(* IEC 61131-3 sources: volt/packages/volt-lsp-iec/test-corpus/awa-palletizer/Device/Plc Logic/Application/Library Manager/L_IPAP_ParameterManagerAccess, 29 files *)

(* ---- L_IPAP_DATATYPE.dut ---- *)
TYPE L_IPAP_DATATYPE :
(
	DT_EMPTY := 0,
	DT_STRING := 1,
	DT_WSTRING := 2,
	DT_BOOLEAN := 3,
	DT_INTEGER_8 := 4,
	DT_INTEGER_16 := 5,
	DT_INTEGER_32 := 6,
	DT_INTEGER_64 := 7,
	DT_UNSIGNED_8 := 8,
	DT_UNSIGNED_16 := 9,
	DT_UNSIGNED_32 := 10,
	DT_UNSIGNED_64 := 11,
	DT_FLOAT_32 := 12,
	DT_FLOAT_64 := 13,
	DT_OCTETSTRING := 14
);
END_TYPE

(* ---- L_IPAP_ERRORID.dut ---- *)
TYPE L_IPAP_ERRORID :
(
	ERR_NOERROR := 0,
	ERR_PARAMETERERROR,
	ERR_INTERNALERROR,
	ERR_TIMEOUT,
	ERR_PARAMETERNOTEXISTING,
	ERR_READACCESSDENIED,
	ERR_WRITEACCESSDENIED,
	ERR_VALUESIZEEXCEEDED,
	ERR_LOWLIMITVIOLATION,
	ERR_HIGHLIMITVIOLATION,
	ERR_NOSELECTLISTVALUE,
	ERR_CONTROLLERINHIBIT,
	ERR_BUFFERSIZE,
	ERR_HAPROXYNOTACTIVE,
	ERR_CHANGEHTTPSREDIRECTFAILED
);
END_TYPE

(* ---- L_IPAP_FBSTATE.dut ---- *)
TYPE L_IPAP_FBSTATE :
(
	INIT := 0,
	WAIT,
	START,
	CHECK,
	DONE,
	ERROR,
	ABORT,
	RESET,
	READ,
	WRITE,
	VERIFY
);
END_TYPE

(* ---- L_IPAP_HTTPSREDIRECT.dut ---- *)
TYPE L_IPAP_HTTPSREDIRECT :
(
	DISABLE_HTTPSREDIRECT := 0,
	ENABLE_HTTPSREDIRECT := 1
);
END_TYPE

(* ---- L_IPAP_INTERNALERROR.dut ---- *)
TYPE L_IPAP_INTERNALERROR :
(
	ERR_OK := 16#0,
	ERR_PROTOCOL_TIMEOUT := 16#2,
	ERR_OUT_OF_MEMORY := 16#4,
	ERR_UNSUPPORTED_ACCESS := 16#5,
	ERR_WRITE_ONLY_ENTRY := 16#6,
	ERR_READ_ONLY_ENTRY := 16#7,
	ERR_OBJECT_NOT_EXISTING := 16#8,
	ERR_PARAM_IS_INCOMPATIBLE := 16#B,
	ERR_INTERNAL_DEVICE_INCOMPATIBILITY := 16#C,
	ERR_PARAM_LENGTH_ERROR := 16#E,
	ERR_PARAM_LENGTH_TOO_LONG := 16#F,
	ERR_PARAM_LENGTH_TOO_SHORT := 16#10,
	ERR_SUBINDEX_NOT_EXISTING := 16#11,
	ERR_VALUE_EXCEEDED := 16#12,
	ERR_VALUE_TOO_GREAT := 16#13,
	ERR_VALUE_TOO_SMALL := 16#14,
	ERR_MAX_VALUE_IS_LESS_THAN_MIN_VALUE := 16#15,
	ERR_GENERAL_ERROR := 16#16,
	ERR_DATA_CANNOT_BE_READ_OR_STORED := 16#17,
	ERR_DATA_CANNOT_BE_READ_OR_STORED_BECAUSE_OF_LOCAL_CONTROL := 16#18,
	ERR_DATA_CANNOT_BE_READ_OR_STORED_IN_THIS_STATE := 16#19,
	ERR_SEND_REQUEST_FAILED := 16#50,
	ERR_UNKNOWN_DATATYPE := 16#51,
	ERR_BUFFER_SIZE := 16#52
);
END_TYPE

(* ---- L_IPAP_INTERNALERROR_ABORTCODE.dut ---- *)
TYPE L_IPAP_INTERNALERROR_ABORTCODE :
(
	ABORT_NOERROR := 16#0,
	ABORT_TIMEOUT := 16#5040000,
	ABORT_OUT_OF_MEMORY := 16#5040005,
	ABORT_UNSUPPORTED_ACCESS := 16#6010000,
	ABORT_WRITE_ONLY_ENTRY := 16#6010001,
	ABORT_READ_ONLY_ENTRY := 16#6010002,
	ABORT_OBJECT_NOT_EXISTING := 16#6020000,
	ABORT_PARAM_IS_INCOMPATIBLE := 16#6040043,
	ABORT_INTERNAL_DEVICE_INCOMPATIBILITY := 16#6040047,
	ABORT_PARAM_LENGTH_ERROR := 16#6070010,
	ABORT_PARAM_LENGTH_TOO_LONG := 16#6070012,
	ABORT_PARAM_LENGTH_TOO_SHORT := 16#6070013,
	ABORT_SUBINDEX_NOT_EXISTING := 16#6090011,
	ABORT_VALUE_EXCEEDED := 16#6090030,
	ABORT_VALUE_TOO_GREAT := 16#6090031,
	ABORT_VALUE_TOO_SMALL := 16#6090032,
	ABORT_MAX_VALUE_IS_LESS_THAN_MIN_VALUE := 16#6090036,
	ABORT_GENERAL_ERROR := 16#8000000,
	ABORT_DATA_CANNOT_BE_READ_OR_STORED := 16#8000020,
	ABORT_DATA_CANNOT_BE_READ_OR_STORED_BECAUSE_OF_LOCAL_CONTROL := 16#8000021,
	ABORT_DATA_CANNOT_BE_READ_OR_STORED_IN_THIS_STATE := 16#8000022
);
END_TYPE

(* ---- L_IPAP_INTERNALERROR_OLD.dut ---- *)
TYPE L_IPAP_INTERNALERROR_OLD :
(
	PMA_OK := 0,
	PMA_TOGGLEBITNOTCHANGED := 1,
	PMA_SDOPROTOCOLTIMEOUT := 2,
	PMA_COMMANDSPECIFIERUNKNOWN := 3,
	PMA_OUTOFMEMORY := 4,
	PMA_UNSUPPORTEDACCESS := 5,
	PMA_WRITEONLYENTRY := 6,
	PMA_READONLYENTRY := 7,
	PMA_OBJECTNOTEXISTING := 8,
	PMA_OBJECTCANTBEPDOMAPPED := 9,
	PMA_MAPPEDOBJECTSEXCEEDPDO := 10,
	PMA_PARAMISINCOMPATIBLE := 11,
	PMA_INTERNALDEVICEINCOMPATIBILITY := 12,
	PMA_HARDWAREERROR := 13,
	PMA_PARAMLENGTHERROR := 14,
	PMA_PARAMLENGTHTOOLONG := 15,
	PMA_PARAMLENGTHTOOSHORT := 16,
	PMA_SUBINDEXNOTEXISTING := 17,
	PMA_VALUEEXCEEDED := 18,
	PMA_VALUETOOGREAT := 19,
	PMA_VALUETOOSMALL := 20,
	PMA_MAXVALUEISLESSTHANMINVALUE := 21,
	PMA_GENERALERROR := 22,
	PMA_DATACANNOTBEREADORSTORED := 23,
	PMA_DATACANNOTBEACCESSEDBECAUSEOFLOCALCONTROL := 24,
	PMA_INTHISSTATEDATACANNOTBEREADORSTORED := 25,
	PMA_NOOBJECTDICTIONARYISPRESENT := 26,
	PMA_ENTRYCANTBEWRITTENSI0NOT0 := 27,
	PMA_COMPLETEACCESSNOTSUPPORTEDFFORTHISOBJ := 28,
	PMA_OBJLENGTHEXCEEDSMBXSIZE := 29,
	PMA_OBJMAPPEDTOPDOSDOACCESSBLOCKED := 30,
	PMA_BUFFEROVERFLOW := 33,
	PMA_INVALIDREPLY := 34,
	PMA_UNKNOWNCOMMAND := 35,
	PMA_PARAMETERERROR := 37,
	PMA_REPLYERROR := 38,
	PMA_REPLYTIMEOUT := 39,
	PMA_SERVERQUEUEERROR := 40,
	PMA_PROTOCOLMISMATCH := 41,
	PMA_SENDREQUESTFAILED := 70,
	PMA_UNKNOWNDATATYPE := 71,
	PMA_OTHERERROR := 99
);
END_TYPE

(* ---- L_IPAP_REQUEST_STATE.dut ---- *)
TYPE L_IPAP_REQUEST_STATE :
(
	UNKNOWN := 0,
	ERROR := 1,
	WAIT := 2,
	BUSY := 3,
	DONE := 4
);
END_TYPE

(* ---- GETBOOLEANPROPERTY.pou ---- *)
FUNCTION GETBOOLEANPROPERTY : BOOL
VAR_INPUT
	STKEY : WSTRING;
END_VAR
END_FUNCTION

(* ---- GETCOMPANY.pou ---- *)
FUNCTION GETCOMPANY : WSTRING
END_FUNCTION

(* ---- GETNUMBERPROPERTY.pou ---- *)
FUNCTION GETNUMBERPROPERTY : DINT
VAR_INPUT
	STKEY : WSTRING;
END_VAR
END_FUNCTION

(* ---- GETTEXTPROPERTY.pou ---- *)
FUNCTION GETTEXTPROPERTY : WSTRING
VAR_INPUT
	STKEY : WSTRING;
END_VAR
END_FUNCTION

(* ---- GETTEXTPROPERTY2.pou ---- *)
FUNCTION GETTEXTPROPERTY2 : POINTER TO WSTRING
VAR_INPUT
	STKEY : WSTRING;
END_VAR
END_FUNCTION

(* ---- GETTITLE.pou ---- *)
FUNCTION GETTITLE : WSTRING
END_FUNCTION

(* ---- GETVERSION.pou ---- *)
FUNCTION GETVERSION : VERSION
END_FUNCTION

(* ---- GETVERSIONPROPERTY.pou ---- *)
FUNCTION GETVERSIONPROPERTY : VERSION
VAR_INPUT
	STKEY : WSTRING;
END_VAR
END_FUNCTION

(* ---- L_IPAP_CHECKREADRESULT.pou ---- *)
FUNCTION L_IPAP_CHECKREADRESULT : L_IPAP_REQUEST_STATE
VAR_INPUT
	HREADREQUEST : RTS_IEC_HANDLE;
	PREADBUFFER : POINTER TO BYTE;
	UIBUFFERSIZE : UDINT;
	PREADDATASIZE : POINTER TO UDINT;
	PREADDATATYPE : POINTER TO L_IPAP_DATATYPE;
	PREQUESTRESULT : POINTER TO RTS_IEC_RESULT;
END_VAR
END_FUNCTION

(* ---- L_IPAP_CHECKWRITERESULT.pou ---- *)
FUNCTION L_IPAP_CHECKWRITERESULT : L_IPAP_REQUEST_STATE
VAR_INPUT
	HWRITEREQUEST : RTS_IEC_HANDLE;
	PREQUESTRESULT : POINTER TO RTS_IEC_RESULT;
END_VAR
END_FUNCTION

(* ---- L_IPAP_ERRORHANDLING.pou ---- *)
FUNCTION L_IPAP_ERRORHANDLING : L_IPAP_ERRORID
VAR_INPUT
	EINTERNALERROR : L_IPAP_INTERNALERROR;
END_VAR
END_FUNCTION

(* ---- L_IPAP_SENDREADREQUEST.pou ---- *)
FUNCTION L_IPAP_SENDREADREQUEST : RTS_IEC_HANDLE
VAR_INPUT
	WINDEX : WORD;
	BYSUBINDEX : BYTE;
END_VAR
END_FUNCTION

(* ---- L_IPAP_SENDREADREQUEST_BASEPM.pou ---- *)
FUNCTION L_IPAP_SENDREADREQUEST_BASEPM : RTS_IEC_HANDLE
VAR_INPUT
	WINDEX : WORD;
	BYSUBINDEX : BYTE;
END_VAR
END_FUNCTION

(* ---- L_IPAP_SENDWRITEREQUEST.pou ---- *)
FUNCTION L_IPAP_SENDWRITEREQUEST : RTS_IEC_HANDLE
VAR_INPUT
	WINDEX : WORD;
	BYSUBINDEX : BYTE;
	UIVALUESIZE : UDINT;
	PVALUE : POINTER TO BYTE;
END_VAR
END_FUNCTION

(* ---- L_IPAP_SENDWRITEREQUEST_BASEPM.pou ---- *)
FUNCTION L_IPAP_SENDWRITEREQUEST_BASEPM : RTS_IEC_HANDLE
VAR_INPUT
	WINDEX : WORD;
	BYSUBINDEX : BYTE;
	UIVALUESIZE : UDINT;
	PVALUE : POINTER TO BYTE;
END_VAR
END_FUNCTION

(* ---- L_IPAP_SENDWRITEREQUEST_INTERNAL.pou ---- *)
FUNCTION L_IPAP_SENDWRITEREQUEST_INTERNAL : RTS_IEC_HANDLE
VAR_INPUT
	WINDEX : WORD;
	BYSUBINDEX : BYTE;
	UIVALUESIZE : UDINT;
	PVALUE : POINTER TO BYTE;
END_VAR
END_FUNCTION

(* ---- GLOBALTEXTLIST.pou ---- *)
FUNCTION_BLOCK GLOBALTEXTLIST
VAR
	M_TEXTLISTFILE : STRING(255);
	_STNAMESPACE : STRING;
END_VAR
END_FUNCTION_BLOCK

(* ---- IMAGEPOOL.pou ---- *)
FUNCTION_BLOCK IMAGEPOOL
VAR
	M_STNAMESPACE : STRING(80);
	M_STHELPVARID : STRING;
	M_STHELPVARPATH : STRING(255);
	M_STHELP : STRING;
	M_REGISTERIMAGES : BOOL := TRUE;
END_VAR
END_FUNCTION_BLOCK

METHOD FB_INIT : BOOL
VAR_INPUT
	BINITRETAINS : BOOL;
	BINCOPYCODE : BOOL;
END_VAR
END_METHOD

METHOD FB_REINIT : BOOL
END_METHOD

METHOD FB_EXIT : BOOL
VAR_INPUT
	BINCOPYCODE : BOOL;
END_VAR
END_METHOD

(* ---- L_IPAP_CHANGEHTTPSREDIRECTSETTING4EASYUI.pou ---- *)
FUNCTION_BLOCK L_IPAP_CHANGEHTTPSREDIRECTSETTING4EASYUI
VAR_INPUT
	XEXECUTE : BOOL;
	XABORT : BOOL;
	EHTTPSREDIRECTSETTING : L_IPAP_HTTPSREDIRECT;
	UDITIMEOUT : UDINT := 0;
END_VAR
VAR_OUTPUT
	XDONE : BOOL;
	XBUSY : BOOL;
	XABORTED : BOOL;
	XERROR : BOOL;
	EERRORID : L_IPAP_ERRORID;
END_VAR
VAR
	FB_TIMEOUT : TON;
	XEXECUTELAST : BOOL;
	XABORTLAST : BOOL;
	BRESETOUTPUT : BOOL;
	BFALLINGEXECUTE : BOOL;
	BFALLINGABORT : BOOL;
	FBSTATE : L_IPAP_FBSTATE;
	MINDEX : WORD;
	MSUBINDEX : BYTE;
	MSETTING : L_IPAP_HTTPSREDIRECT;
	MREQUESTHANDLE : RTS_IEC_HANDLE;
	MREQUESTSTATE : L_IPAP_REQUEST_STATE;
	MREQUESTRESULT : L_IPAP_INTERNALERROR;
	CURSETTING : USINT;
	UDIDATAREAD : UDINT;
	EDATATYPE : L_IPAP_DATATYPE;
END_VAR
END_FUNCTION_BLOCK

(* ---- L_IPAP_PARAMETERREAD.pou ---- *)
FUNCTION_BLOCK L_IPAP_PARAMETERREAD
VAR_INPUT
	XEXECUTE : BOOL;
	XABORT : BOOL;
	XBASEPARAMETER : BOOL := FALSE;
	WINDEX : WORD;
	BYSUBINDEX : BYTE;
	UDITIMEOUT : UDINT := 0;
	PDATABUFFER : POINTER TO BYTE := 0;
	UDIBUFFERSIZE : UDINT := 0;
END_VAR
VAR_OUTPUT
	XDONE : BOOL;
	XBUSY : BOOL;
	XABORTED : BOOL;
	XERROR : BOOL;
	EERRORID : L_IPAP_ERRORID;
	UDIDATAREAD : UDINT;
	EDATATYPE : L_IPAP_DATATYPE;
END_VAR
VAR
	FB_TIMEOUT : TON;
	XEXECUTELAST : BOOL;
	XABORTLAST : BOOL;
	BRESETOUTPUT : BOOL;
	BFALLINGEXECUTE : BOOL;
	BFALLINGABORT : BOOL;
	FBSTATE : L_IPAP_FBSTATE;
	MREQUESTHANDLE : RTS_IEC_HANDLE;
	MREQUESTSTATE : L_IPAP_REQUEST_STATE;
	MREQUESTRESULT : L_IPAP_INTERNALERROR;
END_VAR
END_FUNCTION_BLOCK

(* ---- L_IPAP_PARAMETERWRITE.pou ---- *)
FUNCTION_BLOCK L_IPAP_PARAMETERWRITE
VAR_INPUT
	XEXECUTE : BOOL;
	XABORT : BOOL;
	XBASEPARAMETER : BOOL := FALSE;
	WINDEX : WORD;
	BYSUBINDEX : BYTE;
	UDITIMEOUT : UDINT := 0;
	PDATABUFFER : POINTER TO BYTE := 0;
	UDIDATASIZE : UDINT := 0;
END_VAR
VAR_OUTPUT
	XDONE : BOOL;
	XBUSY : BOOL;
	XABORTED : BOOL;
	XERROR : BOOL;
	EERRORID : L_IPAP_ERRORID;
END_VAR
VAR
	FB_TIMEOUT : TON;
	XEXECUTELAST : BOOL;
	XABORTLAST : BOOL;
	BRESETOUTPUT : BOOL;
	BFALLINGEXECUTE : BOOL;
	BFALLINGABORT : BOOL;
	FBSTATE : L_IPAP_FBSTATE;
	MREQUESTHANDLE : RTS_IEC_HANDLE;
	MREQUESTSTATE : L_IPAP_REQUEST_STATE;
	MREQUESTRESULT : L_IPAP_INTERNALERROR;
END_VAR
END_FUNCTION_BLOCK
